FUNCTION_BLOCK FB_RefMarkerSearch
VAR_INPUT
	Enable					: BOOL;
END_VAR
VAR_OUTPUT
END_VAR
VAR
	Axis						: AXIS_REF;
	Trigger						: TRIGGER_REF;
	bReady	: BOOL;
	btest : Bool;
	Axis_Status:	MC_ReadStatus;
	Axis_Home:		MC_Home;
	Axis_Power:		MC_Power;
	TouchProbe:		MC_TouchProbe;
	
	aRefPoints  : ARRAY [0..100] OF LREAL;
	aDistance	: ARRAY [1..100] OF LREAL;
	nIndx : UINT := 0;
	nState : UINT := 0;
	
	iErrorId					: UDINT;
	iCommandAborted				: BOOL;
END_VAR

// query the status of the axis at the beginning of the cycle
Axis_Status(Enable := TRUE,
			Axis := Axis);

// Enable the axis (power signal or manual enable)
Axis_Power(
	Axis := Axis,
	Enable := Enable,
	Enable_Positive := Enable,
	Enable_Negative := Enable,
	Override := 100.0,
	Status => bReady);

Trigger.EncoderID := 1;
Trigger.Edge := E_SignalEdge.RisingEdge;
Trigger.Mode := E_TouchProbeMode.TOUCHPROBEMODE_SINGLE_COMPATIBILITYMODE;
Trigger.TouchProbe := E_TouchProbe.TouchProbe1;
CASE nState OF
	0 :	(* init *)
		IF bReady AND btest THEN
			nIndx := 0; // reset index
			nState := nState + 1;
		END_IF
		
	1:
		TouchProbe(
			Execute 		:= TRUE,
			Axis 			:= Axis,
			TriggerInput 	:= Trigger,
			RecordedPosition => aRefPoints[nIndx]);
			
		IF NOT TouchProbe.Busy AND TouchProbe.Done THEN
			TouchProbe(	
				Execute			:= FALSE,
				TriggerInput 	:= Trigger, 
				Axis			:= Axis);
			IF nIndx > 0 THEN
				aDistance[nIndx] := F_RoundLREAL(ABS(aRefPoints[nIndx] - aRefPoints[nIndx-1]), 2);
			END_IF
			nIndx := nIndx + 1;
			nState :=  1; 	(* search for next position *)
		ELSIF NOT TouchProbe.Busy AND (TouchProbe.Error OR TouchProbe.CommandAborted) THEN
			iErrorID := TouchProbe.ErrorID;
			
			TouchProbe(	
				Execute			:= FALSE, 
				TriggerInput 	:= Trigger,
				Axis			:= Axis);

			nState 	:= 20;
		END_IF
END_CASE

END_FUNCTION_BLOCK

(* stored: Version 1.1.0.1, ProductVersion 3.1.4024.15
   POU FB_RefMarkerSearch: Id {55946a12-3aba-4836-8e63-10bca96d8d7c}, SpecialFunc None *)
